{attribute 'qualified_only'}
{attribute 'strict'}
{attribute 'to_string'}
TYPE E_AxisReferenceMode : (
    Unknown := 0,
    Incremental := 1,
    Absolute := 2
);
END_TYPE

(* stored: Version 1.1.0.1, ProductVersion 3.1.4026.20
   DUT E_AxisReferenceMode: Id {d18553e8-3b89-54e8-85ca-487a24559bd8} *)
